Fanuc KAREL source: ka00205.KL

PROGRAM KA00205
%STACKSIZE=65535
%PRIORITY=65535
%NOLOCKGROUP
VAR
SRC : ARRAY[4] OF VECTOR
DST : ARRAY[4] OF VECTOR
BEGIN
-- UNRESOLVED_PC line 7 opcodes [22 22 1E] marker_code=0
END KA00205
